//---------------------------------------------------------------------------------------------------------------
//
//  HAUD 2025.12.30
//
//  - fb_ProcessConductor
//  -----------------------------
//  - detects new entry in the cyclic linked list wrapper
//    - forwards the received entry to target instance
//
//  - Ctrl / State for you to use (uses instance ctrl/state pair)
//  - this conductor has no transport process
//  - this conductor is used for sending tickets to a transport process list
//---------------------------------------------------------------------------------------------------------------
FUNCTION_BLOCK fb_ProcessConductor
VAR
  _nConductor             : E_INSTANCE := E_INSTANCE.INSTANCE_CONDUCTOR; // msg device identifier, in case you instantiate more than one conductor
  _stCtrl                 : REFERENCE TO ST_INSTANCE_CTRL;
  _stState                : REFERENCE TO ST_INSTANCE_STATE;

  _eCmd,
  _eCmdOld                : E_INSTANCE_CMD;       // commands for local state machine
  _eStateInstance         : E_INSTANCE_STATE;     // local state machine for infeed procedure

  _eResult                : E_PROGRESS;           // result for methods
  _eStateProgress         : E_PROGRESS;           // substate for local state machine

  _eInit                  : E_PROGRESS;           // startup
  _eCheck                 : E_INSTANCE_CHECK;     // pointer checks

  // the outboxes
  _ItfProcessList         : ARRAY[1..MAX_PROCESS] OF I_Process_LinkedList;  // access to all linked lists for writing tickets
  _WriteResult            : ST_PROCESS_LIST_RESULT;   // last job written to target

  // the inbox
  _ItfTicketList          : I_Process_LinkedList;
  _ResultTicketList       : ST_PROCESS_LIST_RESULT;   // internal list results
  _DeleteResult           : ST_PROCESS_LIST_RESULT;   // last job executed

  _stProcessData          : ST_PROCESS_DATA;          // process target AND station mask

  _stMsg                  : ST_Message;
  _MessageLevel           : E_MessageType := E_MessageType.eMessageInfo;
END_VAR

//-----------------------------------------------------------------------------
//-----------------------------------------------------------------------------
// check pointer and interface
// set message device identification
//-----------------------------------------------------------------------------
IF NOT Check() THEN 
  RETURN; 
END_IF
//-----------------------------------------------------------------------------
// check command
//-----------------------------------------------------------------------------
_eCmd                                         := _stCtrl.Cmd;
IF (_eCmd <> _eCmdOld)
THEN
  CASE _eCmd
  OF
    E_INSTANCE_CMD.INIT:
      _eStateInstance                         := E_INSTANCE_STATE.NULL;
      _eStateProgress                         := E_PROGRESS.PROGRESS_INIT;
  END_CASE
  CmdLog();
  _eCmdOld                                    := _eCmd;
END_IF
//-----------------------------------------------------------------------------
//-----------------------------------------------------------------------------
// state machine for ProcessConductor work
//-----------------------------------------------------------------------------
CASE _eStateInstance
OF
  E_INSTANCE_STATE.NULL:
    // first cycle startup
    _eInit                                    := E_PROGRESS.PROGRESS_INVALID;
    _eStateProgress                           := E_PROGRESS.PROGRESS_INIT;
    _eStateInstance                           := E_INSTANCE_STATE.INIT;


  E_INSTANCE_STATE.INIT:
    //-------------------------------------------------------------------------
    CASE _eStateProgress
    OF
    // E_INSTANCE_STATE.INIT:
    //-------------------------------------------------------------------------
      E_PROGRESS.PROGRESS_INIT:
        IF (_ItfTicketList <> 0)
        THEN
          _eStateProgress                     := E_PROGRESS.PROGRESS_BUSY;
        END_IF
    // E_INSTANCE_STATE.INIT:
    //-------------------------------------------------------------------------
      E_PROGRESS.PROGRESS_BUSY:
        IF _ItfTicketList.InitList()
        THEN
          _eInit                              := E_PROGRESS.PROGRESS_DONE;

          _eStateInstance                     := E_INSTANCE_STATE.DISABLED;
          _eStateProgress                     := E_PROGRESS.PROGRESS_BUSY;
        ELSE
          _eStateProgress                     := E_PROGRESS.PROGRESS_ERROR;
        END_IF
      END_CASE
END_CASE
//-----------------------------------------------------------------------------
// DISABLED:
//  - clear local list result data
//  - wait for enable from the outside
//-----------------------------------------------------------------------------
CASE _eStateInstance
OF
  E_INSTANCE_STATE.DISABLED:
    //-------------------------------------------------------------------------
    CASE _eStateProgress
    OF
      E_PROGRESS.PROGRESS_BUSY:
        CASE _eCmd
        OF
          E_INSTANCE_CMD.ENABLE:              // turn it on!!
            _eStateInstance                   := E_INSTANCE_STATE.DETECTION;
            _eStateProgress                   := E_PROGRESS.PROGRESS_BUSY;
  
            IF (_MessageLevel > E_MessageType.eMessageInfo)
            THEN
              _stMsg.eType                    := E_MessageType.eMessageVerbose;
              _stMsg.eSubdevice               := e_Subdevice.Instance_ProcessConductor;
              _stMsg.iErrorNumber             := 0;
              _stMsg.sText                    := concat(TO_STRING(_eStateInstance), ': ');
              _stMsg.sText                    := concat(_stMsg.sText, TO_STRING(_eStateProgress));
              f_MessageSet(_stMsg);
            END_IF
        END_CASE
    END_CASE
END_CASE
//-----------------------------------------------------------------------------
// DETECTION: 
//  - check inked list and GetHead()
//  - copy job data
//  - switch on process
//-----------------------------------------------------------------------------
CASE _eStateInstance
OF
  E_INSTANCE_STATE.DETECTION:
    //-------------------------------------------------------------------------
    CASE _eStateProgress
    OF
      E_PROGRESS.PROGRESS_BUSY:
        IF (_eCmd = E_INSTANCE_CMD.DISABLE)
        THEN
          _eStateInstance                     := E_INSTANCE_STATE.DISABLED;
          _eStateProgress                     := E_PROGRESS.PROGRESS_BUSY;
  
        ELSIF (_ItfTicketList.Count > 0)
        THEN
          // get new job order for my process
          // the list results carries information about who and where
          _ResultTicketList                   := _ItfTicketList.GetHead();
  
          IF (_ResultTicketList.wState <> 0)
          THEN
            // error in list results must not appear
            // if you land here, there is somethng wrong with the initialization or configuration of the linked list
            _eStateProgress                   := E_PROGRESS.PROGRESS_ERROR;
  
            _stMsg.eType                      := E_MessageType.eMessageError;
            _stMsg.eSubdevice                 := e_Subdevice.Instance_ProcessConductor;
            _stMsg.iErrorNumber               := _ResultTicketList.wState;
            _stMsg.sText                      := concat(TO_STRING(_eStateInstance), ': _ResultTicketList.wState: ');
            _stMsg.sText                      := concat(_stMsg.sText, TO_STRING(_eStateProgress));
            f_MessageSet(_stMsg);
  
          ELSE
            IF (_MessageLevel > E_MessageType.eMessageError)
            THEN
              _stMsg.eType                    := E_MessageType.eMessageInfo;
              _stMsg.eSubdevice               := e_Subdevice.Instance_ProcessConductor;
              _stMsg.iErrorNumber             := _ResultTicketList.stData.wTarget;
              _stMsg.sText                    := concat(TO_STRING(_eStateInstance), ': ');
              _stMsg.sText                    := concat(_stMsg.sText, '_ResultTicketList.stData.wTarget: ');
              _stMsg.sText                    := concat(_stMsg.sText, BitsToString(_ResultTicketList.stData.wTarget));
              f_MessageSet(_stMsg);
            END_IF
  
              // list result contains data for target process
            _stProcessData                    := _ResultTicketList.stData;
  
            IF (_stProcessData.wTarget > 0)
            THEN
              _eStateProgress                 := E_PROGRESS.PROGRESS_PREPARE;
  
  
              IF (_MessageLevel > E_MessageType.eMessageEmpty)
              THEN
                _stMsg.eType                  := E_MessageType.eMessageBatch;
                _stMsg.eSubdevice             := e_Subdevice.Instance_ProcessConductor;
                _stMsg.iErrorNumber           := _stProcessData.nTargetId;
                _stMsg.sText                  := concat(TO_STRING(_eStateProgress), ': ');
                _stMsg.sText                  := concat(_stMsg.sText, TO_STRING(e_message_batch.MSG_BATCH_JOB_STARTED));
                f_MessageSet(_stMsg);
              END_IF
            ELSE
              _ResultTicketList               := _ItfTicketList.RemoveHeadValue();

              IF (_ResultTicketList.wState <> 0)
              THEN
                _stMsg.eType                  := E_MessageType.eMessageError;
                _stMsg.eSubdevice             := e_Subdevice.Instance_ProcessConductor;
                _stMsg.iErrorNumber           := _ResultTicketList.wState;
                _stMsg.sText                  := concat(TO_STRING(_eStateProgress), ': _ResultTicketList.wState: ');
                _stMsg.sText                  := concat(_stMsg.sText, BitsToString(_ResultTicketList.wState));
                f_MessageSet(_stMsg);

                _eStateProgress               := E_PROGRESS.PROGRESS_ERROR;
              END_IF
            END_IF
  
            // check target mask for entries
            IF NOT (_stProcessData.wTarget > 0)
            THEN
              _stMsg.eType                    := E_MessageType.eMessageWarning;
              _stMsg.eSubdevice               := e_Subdevice.Process_LinkedList_CheckData;
              _stMsg.iErrorNumber             := 666;
              _stMsg.sText                    := concat(TO_STRING(_eStateInstance), ': ');
              _stMsg.sText                    := concat(_stMsg.sText, '_ProcessData.wTarget: ');
              _stMsg.sText                    := concat(_stMsg.sText, BitsToString(_stProcessData.wTarget));
              f_MessageSet(_stMsg);
            END_IF
          END_IF
        END_IF
    END_CASE
    CASE _eStateProgress
    OF
      E_PROGRESS.PROGRESS_PREPARE:
        // check process target plausibility
        IF NOT (_stProcessData.nProcessId > 0) OR
           NOT (_stProcessData.nProcessId < E_INSTANCE.INSTANCE_MAX)
        THEN
          _ResultTicketList                   := _ItfTicketList.RemoveHeadValue();
  
          IF (_ResultTicketList.wState <> 0)
          THEN
            _stMsg.eType                      := E_MessageType.eMessageError;
            _stMsg.eSubdevice                 := e_Subdevice.Instance_ProcessConductor;
            _stMsg.iErrorNumber               := _ResultTicketList.wState;
            _stMsg.sText                      := concat(TO_STRING(_eStateProgress), ': _ResultTicketList.wState: ');
            _stMsg.sText                      := concat(_stMsg.sText, BitsToString(_ResultTicketList.wState));
            f_MessageSet(_stMsg);

            _eStateProgress                   := E_PROGRESS.PROGRESS_ERROR;
          END_IF

          _stMsg.eType                        := E_MessageType.eMessageError;
          _stMsg.eSubdevice                   := e_Subdevice.Process_LinkedList_CheckData;
          _stMsg.iErrorNumber                 := 6666;
          _stMsg.sText                        := concat(TO_STRING(_eStateInstance), ': ');
          _stMsg.sText                        := concat(_stMsg.sText, '_stProcessData.nProcessId: ');
          _stMsg.sText                        := concat(_stMsg.sText, TO_STRING(_stProcessData.nProcessId));
          f_MessageSet(_stMsg);
  
        ELSE
          IF (_MessageLevel > E_MessageType.eMessageInfo)
          THEN
            _stMsg.eType                      := E_MessageType.eMessageVerbose;
            _stMsg.eSubdevice                 := e_Subdevice.Instance_ProcessConductor;
            _stMsg.iErrorNumber               := _stProcessData.nProcessId;
            _stMsg.sText                      := concat(TO_STRING(_eStateInstance), ': _stProcessData.nProcessId: ');
            _stMsg.sText                      := concat(_stMsg.sText, TO_STRING(_stProcessData.nProcessId));
            f_MessageSet(_stMsg);
          END_IF
  
          _DeleteResult                       := _ItfTicketList.RemoveHeadValue();
  
          IF (_DeleteResult.wState = 0)
          THEN
            _eStateInstance                   := E_INSTANCE_STATE.WORKING;
            _eStateProgress                   := E_PROGRESS.PROGRESS_BUSY;
          ELSE
            _stMsg.eType                      := E_MessageType.eMessageError;
            _stMsg.eSubdevice                 := e_Subdevice.Instance_ProcessConductor;
            _stMsg.iErrorNumber               := _DeleteResult.wState;
            _stMsg.sText                      := concat(TO_STRING(_eStateProgress), ': _DeleteResult.wState: ');
            _stMsg.sText                      := concat(_stMsg.sText, BitsToString(_DeleteResult.wState));
            f_MessageSet(_stMsg);

            _eStateProgress                   := E_PROGRESS.PROGRESS_ERROR;
          END_IF
        END_IF
    END_CASE
END_CASE
//-----------------------------------------------------------------------------
// WORKING
//  - Add ticket in target list
//  - check and log
//  - transition to finish
//-----------------------------------------------------------------------------
CASE _eStateInstance
OF
  E_INSTANCE_STATE.WORKING:
    //-------------------------------------------------------------------------
    CASE _eStateProgress
    OF
      E_PROGRESS.PROGRESS_BUSY:
        // write process ticket, then go back up
        _WriteResult                          := _ItfProcessList[_stProcessData.nProcessId].AddTailValue(_stProcessData);

        IF (_WriteResult.wState <> 0)
        THEN
          // adding to target list must be successful on the first try
          // IF you land here, there is something wrong with initialization or configuration of the linked list
          _stMsg.eType                        := E_MessageType.eMessageError;
          _stMsg.eSubdevice                   := e_Subdevice.Instance_ProcessConductor;
          _stMsg.iErrorNumber                 := _WriteResult.wState;
          _stMsg.sText                        := concat(TO_STRING(_eStateProgress), ': _WriteResult.wState: ');
          _stMsg.sText                        := concat(_stMsg.sText, BitsToString(_WriteResult.wState));
          f_MessageSet(_stMsg);

          _eStateProgress                     := E_PROGRESS.PROGRESS_ERROR;

        ELSE
          _eStateInstance                     := E_INSTANCE_STATE.FINISH;
          _eStateProgress                     := E_PROGRESS.PROGRESS_BUSY;

          IF (_MessageLevel > E_MessageType.eMessageError)
          THEN
            _stMsg.eType                      := E_MessageType.eMessageInfo;
            _stMsg.eSubdevice                 := e_Subdevice.Process_LinkedList_AddTail;
            _stMsg.iErrorNumber               := _stProcessData.nProcessId;
            _stMsg.sText                      := concat(TO_STRING(_eStateInstance), ': _stProcessData.nProcessId: ');
            _stMsg.sText                      := concat(_stMsg.sText, TO_STRING(_stProcessData.nProcessId));

            f_MessageSet(_stMsg);
          END_IF
        END_IF
    END_CASE
END_CASE
//-----------------------------------------------------------------------------
// FINISH:
//-----------------------------------------------------------------------------
CASE _eStateInstance
OF
  E_INSTANCE_STATE.FINISH:
    //-------------------------------------------------------------------------
    CASE _eStateProgress
    OF
      E_PROGRESS.PROGRESS_BUSY:
        _eStateProgress                       := E_PROGRESS.PROGRESS_DONE;
    END_CASE
    // E_INSTANCE_STATE.FINISH:
    //-------------------------------------------------------------------------
    CASE _eStateProgress
    OF
      E_PROGRESS.PROGRESS_DONE:
        _eStateInstance                       := E_INSTANCE_STATE.DISABLED;
        _eStateProgress                       := E_PROGRESS.PROGRESS_BUSY;

    END_CASE
END_CASE
//-----------------------------------------------------------------------------
//-----------------------------------------------------------------------------
_stState.ProcessIdentity                      := _nConductor;
_stState.ProcessState                         := _eStateInstance;
_stState.ProcessProgress                      := _eStateProgress;
_stState.QueueProcessCount                    := TO_UINT(_ItfTicketList.Count);
//-----------------------------------------------------------------------------
//-----------------------------------------------------------------------------

METHOD PUBLIC BitGet : BOOL
VAR_INPUT
  inVal   : T_PROCESS;
  bitNo   : DINT;
END_VAR
VAR
  wConst : T_PROCESS := 1;
END_VAR
IF ( inVal AND SHL( wConst,TO_SINT(bitNo) MOD TO_INT(SIZEOF(T_PROCESS)*8) ) ) > 0
THEN
  BitGet := TRUE;
ELSE
  BitGet := FALSE;
END_IF
END_METHOD

METHOD BitsToString : STRING(SIZEOF(T_PROCESS)*8) // T_PROCESS to string
VAR_INPUT
  inVal       : T_PROCESS;
END_VAR
VAR
  _nx         : DINT;
  _str        : STRING(SIZEOF(T_PROCESS)*8);
END_VAR
FOR _nx := ((SIZEOF(inVal)*8)) TO 1 BY(-1)
DO
  IF (BitGet(inVal, _nx-1))
  THEN
    _str     := concat(_str, '1');
  ELSE
    _str     := concat(_str, '0');
  END_IF
END_FOR

BitsToString := _str;
END_METHOD

METHOD Check  : BOOL // call this method in the extending/inheriting class
VAR_INST
  _idx        : UINT;
END_VAR
//-----------------------------------------------------------------------------
//-----------------------------------------------------------------------------
// pointer checks
//-----------------------------------------------------------------------------
IF NOT __ISVALIDREF(_stCtrl)
THEN
  _eCheck                 := E_INSTANCE_CHECK.INVALID_INSTANCE_CONTROL_REFERENCE;
  RETURN;
END_IF

IF NOT __ISVALIDREF(_stState)
THEN
  _eCheck                 := E_INSTANCE_CHECK.INVALID_INSTANCE_STATE_REFERENCE;
  RETURN;
END_IF

FOR _idx := 1 TO MAX_PROCESS
DO
  IF NOT (_ItfProcessList[_idx] <> 0)
  THEN
    _eCheck               := E_INSTANCE_CHECK.PROCESS_LIST_ITF_INDEX_INVALID;
    RETURN;
  END_IF
END_FOR

IF NOT (_ItfTicketList <> 0)
THEN
  _eCheck                 := E_INSTANCE_CHECK.TICKET_LIST_ITF_INVALID;
  RETURN;
END_IF

//-----------------------------------------------------------------------------
//-----------------------------------------------------------------------------
// set message device
//-----------------------------------------------------------------------------
_stMsg.eDevice            := e_Device.Conductor + TO_UINT(_nConductor);
//-----------------------------------------------------------------------------
//-----------------------------------------------------------------------------
_eCheck                   := E_INSTANCE_CHECK.CHECK_DONE;
Check                     := TRUE;
END_METHOD

METHOD CmdLog

IF (_MessageLevel > E_MessageType.eMessageError)
THEN
  _stMsg.eSubdevice       := e_Subdevice.Instance_ProcessConductor;
  _stMsg.iErrorNumber     := 0;
  _stMsg.sText            := concat('E_INSTANCE_CMD', '.');
  _stMsg.sText            := concat(_stMsg.sText, TO_STRING(_eCmd));
  f_MessageSet(_stMsg);
END_IF
END_METHOD

PROPERTY Ctrl : REFERENCE TO ST_INSTANCE_CTRL
SET
_stCtrl ref= Ctrl;
END_SET
END_PROPERTY

PROPERTY MessageLevel : e_MessageType
GET
MessageLevel := _MessageLevel;
END_GET
SET
_MessageLevel := MessageLevel;
END_SET
END_PROPERTY

PROPERTY ProcessLinkedLists : ARRAY[1..max_process] OF I_Process_LinkedList
SET
_ItfProcessList := ProcessLinkedLists;
END_SET
END_PROPERTY

PROPERTY State : REFERENCE TO ST_INSTANCE_STATE
SET
_stState ref= State;
END_SET
END_PROPERTY

PROPERTY TicketLinkedList : I_Process_LinkedList
SET
_ItfTicketList := TicketLinkedList;
END_SET
END_PROPERTY

END_FUNCTION_BLOCK

(* stored: Version 1.1.0.1, ProductVersion 3.1.4026.20
   POU fb_ProcessConductor: Id {f1a261a4-f63d-4608-955f-a4e7d0d9bbab}, SpecialFunc None
   Method BitGet: Id {2ba1ed32-cb22-46cd-9284-cb807e052273}
   Method BitsToString: Id {56309c51-f8d0-4b4d-ba61-91c4c72e022c}
   Method Check: Id {02cef509-b143-447b-84a9-3ff41a696353}
   Method CmdLog: Id {e5a4e297-c28d-45b7-9a6e-7f0812358825}
   Property Ctrl: Id {be4943df-b340-4c7d-b3b7-947b1d9c86ca}
   Set Set: Id {fb203d93-59c2-4994-815a-f3a55423f261}
   Property MessageLevel: Id {6b37c0b1-2a95-468d-8dc2-6917b103df06}
   Get Get: Id {ebb30769-0926-4ec7-ab5a-6c1a0d486240}
   Set Set: Id {556216a4-55f5-4288-886c-344557b07d7a}
   Property ProcessLinkedLists: Id {3c662d17-f90d-4398-9000-5b26b6e3edad}
   Set Set: Id {3f745bf3-f708-4f4b-8b09-c42abf62b996}
   Property State: Id {b62ba3c2-e868-4e5c-8b87-05f191f1e974}
   Set Set: Id {2154d7fa-134c-4ee1-88b3-077d1ea5ea3c}
   Property TicketLinkedList: Id {282b2c15-5056-4260-97c1-e721960266b4}
   Set Set: Id {278204fe-1707-4511-9bfd-b8b81dec9fb8} *)
